Fanuc KAREL source: kt00743.KL

-- PROVISIONAL review KL for V770-1; original PC SHA256 a0ee91a0cc4bb0e7775c6787aaa3ad5a66c9ff8ceb27c68006dcf868a12472ec
-- Incomplete behavior may be omitted. Consult companion uncertainty JSON. Do not deploy.
PROGRAM KT00743
%NOLOCKGROUP
VAR
  OUT : INTEGER
-- UNRESOLVED_DECL ARG type=002013
BEGIN
  -- UNRESOLVED_PC offsets 5-18; opcodes 22,1D,23
  -- UNRESOLVED_PC offsets 23-27; opcodes 7F
END KT00743
